(* PLC project Unnamed, Unknown Unnamed 1 *)
(* stored: creationDateTime 2026-11-16T11:19:02, modificationDateTime 2026-11-16T11:19:02 *)

FUNCTION_BLOCK TON
  VAR_OUTPUT
    Q : BOOL;
    ET : TIME;
  END_VAR
  VAR_INPUT
    IN : BOOL;
    PT : TIME;
  END_VAR

END_FUNCTION_BLOCK

FUNCTION_BLOCK PRODUCT_SIMULATOR
  VAR
    ARRIVAL_TIMER : TON;
    RANDOM_SEED : DINT := 12345;
    RANDOM_VALUE : DINT := 0;
    SIM_STATE : INT := 0;
    CLEAR_TIMER : TON;
  END_VAR
  VAR_INPUT
    READY : BOOL;
    CONVEYOR : BOOL;
    ACCEPTED : BOOL;
    REJECTED : BOOL;
    REJECTING : BOOL;
    PACKAGING : BOOL;
    TARGET_REACHED : BOOL;
    DEFECT_RATE : INT;
  END_VAR
  VAR_OUTPUT
    SENSOR_OUT : BOOL;
    QUALITY_OUT : BOOL;
  END_VAR

            (* Virtual product arrival timer *)
ARRIVAL_TIMER(
    IN := READY AND CONVEYOR
          AND NOT TARGET_REACHED
          AND (SIM_STATE = 0),
    PT := T#2s
);

(* Product clearance delay *)
CLEAR_TIMER(
    IN := SIM_STATE = 30,
    PT := T#1s
);

IF NOT READY THEN

    SENSOR_OUT := FALSE;
    QUALITY_OUT := FALSE;
    SIM_STATE := 0;

ELSE

    CASE SIM_STATE OF

        0:
            (* Wait for next product *)
            IF ARRIVAL_TIMER.Q THEN
                SIM_STATE := 10;
            END_IF;

        10:
            (* Generate pseudorandom quality *)
            RANDOM_SEED :=
                (RANDOM_SEED * 25173 + 13849)
                MOD 65536;

            RANDOM_VALUE :=
                (RANDOM_SEED * 100) / 65536;

            QUALITY_OUT :=
                RANDOM_VALUE <
                INT_TO_DINT(DEFECT_RATE);

            SENSOR_OUT := TRUE;
            SIM_STATE := 20;

        20:
            (* Wait until product is finished *)
            IF ACCEPTED AND NOT PACKAGING THEN

                SIM_STATE := 30;

            ELSIF REJECTED AND NOT REJECTING THEN

                SIM_STATE := 30;

            END_IF;

        30:
            (* Clear simulated product *)
            SENSOR_OUT := FALSE;

            IF CLEAR_TIMER.Q THEN
                QUALITY_OUT := FALSE;
                SIM_STATE := 0;
            END_IF;

    ELSE
        SENSOR_OUT := FALSE;
        QUALITY_OUT := FALSE;
        SIM_STATE := 0;

    END_CASE;

END_IF;
          
END_FUNCTION_BLOCK

FUNCTION ADD : ANY_NUM
  VAR_INPUT
    IN1 : ANY_NUM;
    IN2 : ANY_NUM;
  END_VAR

END_FUNCTION

FUNCTION_BLOCK CTU
  VAR_OUTPUT
    Q : BOOL;
    CV : INT;
  END_VAR
  VAR_INPUT
    CU : BOOL;
    R : BOOL;
    PV : INT;
  END_VAR

END_FUNCTION_BLOCK

FUNCTION GE : BOOL
  VAR_INPUT
    IN1 : ANY_ELEMENTARY;
    IN2 : ANY_ELEMENTARY;
  END_VAR

END_FUNCTION

FUNCTION GT : BOOL
  VAR_INPUT
    IN1 : ANY_ELEMENTARY;
    IN2 : ANY_ELEMENTARY;
  END_VAR

END_FUNCTION

FUNCTION SUB : ANY_NUM
  VAR_INPUT
    IN1 : ANY_NUM;
    IN2 : ANY_NUM;
  END_VAR

END_FUNCTION

FUNCTION_BLOCK TP
  VAR_OUTPUT
    Q : BOOL;
    ET : TIME;
  END_VAR
  VAR_INPUT
    IN : BOOL;
    PT : TIME;
  END_VAR

END_FUNCTION_BLOCK

PROGRAM main
  VAR
    START AT %QX0.0 : BOOL := FALSE;
    STOP AT %QX0.1 : BOOL := FALSE;
    SYSTEM_RUN AT %QX1.0 : BOOL := FALSE;
    MOTOR AT %QX1.2 : BOOL := FALSE;
    WARNING_LIGHT AT %QX1.1 : BOOL := FALSE;
    PRODUCT_SENSOR AT %QX2.0 : BOOL := FALSE;
    PROCESSOR AT %QX1.3 : BOOL := FALSE;
    INSPECTION_ACTIVE AT %QX1.4 : BOOL := FALSE;
    QUALITY_FAIL AT %QX2.1 : BOOL := FALSE;
    REJECT_ACTIVE AT %QX1.5 : BOOL := FALSE;
    ACCEPT_COUNT AT %QW3 : INT := 0;
    REJECT_COUNT AT %QW4 : INT := 0;
    RESET_COUNTS AT %QX0.2 : BOOL := FALSE;
    TOTAL_PROCESSED AT %QW5 : INT := 0;
    ORDER_QUANTITY AT %QW0 : INT := 20;
    ORDER_REMAINING AT %QW6 : INT := 20;
    ORDER_COMPLETE AT %QX1.7 : BOOL := FALSE;
    BATCH_CAPACITY AT %QW1 : INT := 10;
    BATCH_COUNT AT %QW7 : INT := 0;
    PACKAGE_COUNT AT %QW8 : INT := 0;
    PACKAGING_ACTIVE AT %QX1.6 : BOOL := FALSE;
    DEFECT_PERCENT AT %QW2 : INT := 25;
  END_VAR
  VAR
    STARTUP_TIMER : TON;
    LINE_READY : BOOL := FALSE;
    PROCESS_ACTIVE : BOOL := FALSE;
    PROCESS_DONE : BOOL := FALSE;
    PROCESS_TIMER : TON;
    WAIT_CLEAR : BOOL := FALSE;
    INSPECTION_DONE : BOOL := FALSE;
    INSPECTION_TIMER : TON;
    REJECT_PULSE : BOOL := FALSE;
    PRODUCT_ACCEPTED : BOOL := FALSE;
    PRODUCT_REJECTED : BOOL := FALSE;
    REJECT_TIMER : TP;
    ACCEPT_COUNTER : CTU;
    REJECT_COUNTER : CTU;
    QUANTITY_REACHED : BOOL := FALSE;
    BATCH_COUNTER : CTU;
    PACKAGE_COUNTER : CTU;
    PACKAGING_TIMER : TON;
    BATCH_FULL : BOOL := FALSE;
    BATCH_NOT_READY : BOOL := FALSE;
    PACKAGING_DONE : BOOL := FALSE;
    SIMULATOR : PRODUCT_SIMULATOR;
  END_VAR

(* LD diagram, written out as Structured Text *)
SYSTEM_RUN := NOT STOP AND NOT ORDER_COMPLETE AND (START OR SYSTEM_RUN);
STARTUP_TIMER(IN := SYSTEM_RUN, PT := T#6s);
LINE_READY := STARTUP_TIMER.Q;
WARNING_LIGHT := SYSTEM_RUN AND NOT LINE_READY;
MOTOR := LINE_READY AND NOT PROCESS_ACTIVE AND NOT PRODUCT_SENSOR AND NOT INSPECTION_ACTIVE AND NOT REJECT_ACTIVE AND NOT BATCH_FULL AND NOT PACKAGING_ACTIVE AND NOT QUANTITY_REACHED;
PROCESS_TIMER(IN := LINE_READY AND PROCESS_ACTIVE, PT := T#10s);
PROCESS_DONE := PROCESS_TIMER.Q;
PROCESS_ACTIVE := LINE_READY AND NOT PROCESS_DONE AND NOT WAIT_CLEAR AND NOT INSPECTION_ACTIVE AND NOT REJECT_ACTIVE AND NOT BATCH_FULL AND NOT PACKAGING_ACTIVE AND NOT QUANTITY_REACHED AND (PRODUCT_SENSOR OR PROCESS_ACTIVE);
PROCESSOR := PROCESS_ACTIVE;
WAIT_CLEAR := LINE_READY AND PRODUCT_SENSOR AND (PROCESS_DONE OR WAIT_CLEAR);
INSPECTION_ACTIVE := LINE_READY AND NOT INSPECTION_DONE AND (PROCESS_DONE OR INSPECTION_ACTIVE);
INSPECTION_TIMER(IN := INSPECTION_ACTIVE, PT := T#4s);
INSPECTION_DONE := INSPECTION_TIMER.Q;
IF INSPECTION_DONE AND NOT QUALITY_FAIL THEN PRODUCT_ACCEPTED := TRUE; END_IF;
IF INSPECTION_DONE AND QUALITY_FAIL THEN PRODUCT_REJECTED := TRUE; END_IF;
REJECT_TIMER(IN := PRODUCT_REJECTED, PT := T#1s);
REJECT_PULSE := REJECT_TIMER.Q;
REJECT_ACTIVE := LINE_READY AND REJECT_PULSE;
IF NOT PRODUCT_SENSOR OR NOT LINE_READY THEN PRODUCT_ACCEPTED := FALSE; END_IF;
IF NOT PRODUCT_SENSOR OR NOT LINE_READY THEN PRODUCT_REJECTED := FALSE; END_IF;
QUANTITY_REACHED := ACCEPT_COUNT >= ORDER_QUANTITY;
BATCH_COUNTER(CU := PRODUCT_ACCEPTED, R := PACKAGING_DONE OR RESET_COUNTS, PV := BATCH_CAPACITY);
BATCH_FULL := BATCH_COUNTER.Q;
BATCH_NOT_READY := BATCH_COUNT > 0;
PACKAGING_ACTIVE := LINE_READY AND (BATCH_FULL OR QUANTITY_REACHED AND BATCH_NOT_READY);
PACKAGING_TIMER(IN := PACKAGING_ACTIVE, PT := T#4s);
PACKAGING_DONE := PACKAGING_TIMER.Q;
ORDER_COMPLETE := QUANTITY_REACHED AND NOT BATCH_NOT_READY AND NOT PACKAGING_ACTIVE;
SIMULATOR(READY := LINE_READY, CONVEYOR := MOTOR, ACCEPTED := PRODUCT_ACCEPTED, REJECTED := PRODUCT_REJECTED, REJECTING := REJECT_ACTIVE, PACKAGING := PACKAGING_ACTIVE, TARGET_REACHED := QUANTITY_REACHED, DEFECT_RATE := DEFECT_PERCENT);
PRODUCT_SENSOR := SIMULATOR.SENSOR_OUT;
QUALITY_FAIL := SIMULATOR.QUALITY_OUT;
 := STARTUP_TIMER.ET;
 := PROCESS_TIMER.ET;
 := INSPECTION_TIMER.ET;
 := REJECT_TIMER.ET;
ACCEPT_COUNTER(CU := PRODUCT_ACCEPTED, R := RESET_COUNTS, PV := 32767);
ACCEPT_COUNT := ACCEPT_COUNTER.CV;
REJECT_COUNTER(CU := PRODUCT_REJECTED, R := RESET_COUNTS, PV := 32767);
REJECT_COUNT := REJECT_COUNTER.CV;
TOTAL_PROCESSED := ACCEPT_COUNT + REJECT_COUNT;
ORDER_REMAINING := ORDER_QUANTITY - ACCEPT_COUNT;
BATCH_COUNT := BATCH_COUNTER.CV;
 := PACKAGING_TIMER.ET;
PACKAGE_COUNTER(CU := PACKAGING_DONE, R := RESET_COUNTS, PV := 32767);
PACKAGE_COUNT := PACKAGE_COUNTER.CV;
END_PROGRAM

CONFIGURATION Config0
  RESOURCE Res0 ON PLC
    TASK task0(INTERVAL := T#20ms, PRIORITY := 1);
    PROGRAM instance0 WITH task0 : main;
  END_RESOURCE
END_CONFIGURATION
